(* IEC 61131-3 sources: helmsman/crates/helmsman-canvas/assets/front, 6 files *)

(* ---- main.st ---- *)
PROGRAM tank
VAR_INPUT
  level_low : BOOL;
  level_high : BOOL;
  level : REAL := 1.0;    (* metres, tank is 2 m deep *)
  reset : BOOL;
END_VAR
VAR_OUTPUT
  fill : BOOL;            (* inlet valve *)
  alarm : BOOL;
  level_pct : REAL;       (* level for the operator's screen *)
END_VAR
VAR
  fill_time : TON;        (* how long the inlet has been open *)
  overrun_trip : BOOL;    (* a fill ran past 7 s: inlet shut, alarm up *)
  switches_disagree : BOOL; (* low and high both on: inlet shut, alarm up *)
  alarm_latch : BOOL;     (* alarm held until reset with the switches agreed *)
END_VAR

(* Level readout: 0 m -> 0 %, 2 m -> 100 %. *)
level_pct := LIMIT(0.0, level / 2.0 * 100.0, 100.0);

(* A fill takes under 6 s: one that runs 7 s trips the overrun. *)
fill_time(IN := fill, PT := T#7s);
IF fill_time.Q THEN
  overrun_trip := TRUE;
END_IF;
IF reset THEN
  overrun_trip := FALSE;
END_IF;

(* Both switches on at once: the level cannot be low and full, so
   close the inlet and alarm. *)
switches_disagree := level_low AND level_high;

(* Alarm hold: any cause sets the latch; only reset pressed while the
   switches agree clears it. *)
IF overrun_trip OR switches_disagree THEN
  alarm_latch := TRUE;
END_IF;
IF reset AND NOT switches_disagree THEN
  alarm_latch := FALSE;
END_IF;

(* Top-up: open the inlet when the tank runs low, close it when full,
   when a fill has run too long, when the switches disagree, or while
   the alarm is held. *)
fill := (level_low OR fill) AND NOT level_high
        AND NOT overrun_trip AND NOT switches_disagree
        AND NOT alarm_latch;

alarm := alarm_latch;
END_PROGRAM

(* ---- test_alarm_needs_reset.st ---- *)
(* An alarm stays on, and the inlet closed, until someone presses reset. *)
PROGRAM test_alarm_needs_reset
VAR_INPUT
  fill  : BOOL;
  alarm : BOOL;
END_VAR
VAR_OUTPUT
  level_high_stuck : BOOL;
  reset : BOOL;
  done : BOOL;
END_VAR
VAR
  seen : BOOL;
  after : TON;
  pressed : TON;
  still_on : ASSERT;      (* the alarm stayed on after the fault went away *)
  still_closed : ASSERT;  (* the inlet stayed closed *)
  cleared : ASSERT;       (* reset cleared the alarm *)
END_VAR
(* The high switch fails until the alarm comes on, then works again. *)
IF alarm THEN
  seen := TRUE;
END_IF;
level_high_stuck := NOT seen;
after(IN := seen, PT := T#3s);
IF after.Q AND NOT reset THEN
  still_on(COND := alarm);
  still_closed(COND := NOT fill);
  reset := TRUE;
END_IF;
pressed(IN := reset, PT := T#500ms);
IF pressed.Q THEN
  cleared(COND := NOT alarm);
  done := TRUE;
END_IF;
END_PROGRAM

(* ---- test_both_switches_on.st ---- *)
(* Nearly empty and full at once cannot be true: the inlet stays closed and the alarm comes on. *)
PROGRAM test_both_switches_on
VAR_INPUT
  fill  : BOOL;
  alarm : BOOL;
END_VAR
VAR_OUTPUT
  level_low  : BOOL;
  level_high : BOOL;
  done : BOOL;
END_VAR
VAR
  t : TON;
  inlet_closed : ASSERT;  (* the inlet is closed *)
  alarm_on : ASSERT;      (* the alarm is on *)
END_VAR
level_low := TRUE;
level_high := TRUE;
t(IN := TRUE, PT := T#1s);
IF t.Q THEN
  inlet_closed(COND := NOT fill);
  alarm_on(COND := alarm);
  done := TRUE;
END_IF;
END_PROGRAM

(* ---- test_fills_and_stops.st ---- *)
(* The inlet opens when the tank runs low and closes again when it is full. *)
PROGRAM test_fills_and_stops
VAR_INPUT
  fill  : BOOL;
  alarm : BOOL;
END_VAR
VAR_OUTPUT
  done : BOOL;
END_VAR
VAR
  t : TON;
  opened : BOOL;
  closed_again : BOOL;
  inlet_opened_when_low : ASSERT;   (* the inlet opened when the tank ran low *)
  inlet_closed_when_full : ASSERT;  (* the inlet closed when the tank was full *)
  no_alarm : ASSERT;                (* no alarm in a normal fill *)
END_VAR
t(IN := TRUE, PT := T#20s);
IF fill THEN
  opened := TRUE;
END_IF;
IF opened AND NOT fill THEN
  closed_again := TRUE;
END_IF;
IF t.Q THEN
  inlet_opened_when_low(COND := opened);
  inlet_closed_when_full(COND := closed_again);
  no_alarm(COND := NOT alarm);
  done := TRUE;
END_IF;
END_PROGRAM

(* ---- test_high_switch_fails.st ---- *)
(* If the high switch fails, the inlet still closes before the tank overflows, and the alarm comes on. *)
PROGRAM test_high_switch_fails
VAR_INPUT
  fill  : BOOL;
  alarm : BOOL;
END_VAR
VAR_OUTPUT
  level_high_stuck : BOOL;
  done : BOOL;
END_VAR
VAR
  t : TON;
  overflow : TON;
  overflowed : BOOL;
  inlet_closed : ASSERT;      (* the inlet is closed *)
  alarm_on : ASSERT;          (* the alarm is on *)
  never_overflowed : ASSERT;  (* the inlet was never open long enough to overflow the tank *)
END_VAR
(* The high switch never makes. *)
level_high_stuck := TRUE;
t(IN := TRUE, PT := T#20s);
(* From nearly empty, 7.2 s of filling reaches the brim. *)
overflow(IN := fill, PT := T#7s200ms);
IF overflow.Q THEN
  overflowed := TRUE;
END_IF;
IF t.Q THEN
  inlet_closed(COND := NOT fill);
  alarm_on(COND := alarm);
  never_overflowed(COND := NOT overflowed);
  done := TRUE;
END_IF;
END_PROGRAM

(* ---- test_switches_lost.st ---- *)
(* If the level switches are lost while the tank is filling, the inlet closes. *)
PROGRAM test_switches_lost
VAR_INPUT
  fill : BOOL;
END_VAR
VAR_OUTPUT
  level_low_absent : BOOL;
  done : BOOL;
END_VAR
VAR
  t : TON;
  was_filling : BOOL;
  lost : TON;
  filling_before : ASSERT;  (* the tank was filling when the switches were lost *)
  inlet_closed : ASSERT;    (* the inlet closed *)
END_VAR
t(IN := TRUE, PT := T#4s);
IF fill AND NOT t.Q THEN
  was_filling := TRUE;
END_IF;
(* 4 s in, mid-fill, the module the switches are wired to goes away. *)
level_low_absent := t.Q;
lost(IN := t.Q, PT := T#1s);
IF lost.Q THEN
  filling_before(COND := was_filling);
  inlet_closed(COND := NOT fill);
  done := TRUE;
END_IF;
END_PROGRAM
